FUNCTION_BLOCK MOD_StateManager (* The module's PackML state: Stopped, Resetting, Idle, Execute, Stopping, Aborted. The owner changes it with the OPC UA methods Reset, Start, Stop, Abort and Clear. It runs the Resetting and Stopping procedures and publishes the state for clients and for every block. Technical: Module state manager: OPC UA methods Reset/Start/Stop/Abort/Clear(Session) answer [Accepted, ErrorID]; publishes the PackML State over OPC UA and on the module's state channel; RUN_RESETTING and RUN_STOPPING start the procedures, which answer with *_DONE or *_FAILED *)
  (* Standard: 61499-2 *)
  (* Version 0.1, 2026-09-28, Project contributors, AAU Smart Production Lab *)
  PACKAGE modlib;
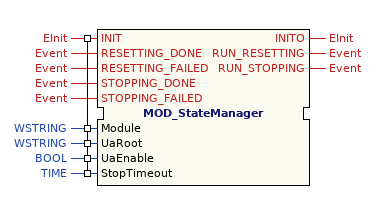
  EVENT_INPUT
    INIT : EInit WITH Module, UaRoot, UaEnable, StopTimeout; (* Initialise, once at start-up (the INIT chain); takes the values given with it *)
    RESETTING_DONE; (* The Resetting procedure ended *)
    RESETTING_FAILED; (* The Resetting procedure failed *)
    STOPPING_DONE; (* The Stopping procedure ended *)
    STOPPING_FAILED; (* The Stopping procedure failed *)
  END_EVENT
  EVENT_OUTPUT
    INITO : EInit; (* Initialised: the next block of the INIT chain goes on *)
    RUN_RESETTING; (* Run the Resetting procedure (the module was reset) *)
    RUN_STOPPING; (* Run the Stopping procedure (the module was stopped) *)
  END_EVENT
  VAR_INPUT
    Module : WSTRING; (* The module's name; its local channels are named after it (loc[<Module>/...]) *)
    UaRoot : WSTRING; (* The module's OPC UA folder, e.g. /Objects/Filling *)
    UaEnable : BOOL; (* Publish on OPC UA *)
    StopTimeout : TIME := T#10s; (* How long Stopping may take before the module aborts *)
  END_VAR
  FBS
    Ids : modlib::MOD_StateIds; (* Builds the OPC UA addresses and channel names from the module's name. *)
    Owner : modlib::MOD_OwnerView; (* Knows who occupies the module: only the owner may change the state. *)
    Reset : iec61499::net::SERVER_2_1; (* The OPC UA method Module/Reset(Session). *)
    Start : iec61499::net::SERVER_2_1; (* The OPC UA method Module/Start(Session). *)
    Stop : iec61499::net::SERVER_2_1; (* The OPC UA method Module/Stop(Session). *)
    Abort : iec61499::net::SERVER_2_1; (* The OPC UA method Module/Abort(Session). *)
    Clear : iec61499::net::SERVER_2_1; (* The OPC UA method Module/Clear(Session). *)
    Gate : modlib::MOD_StateGate; (* Decides the commands: only from the owner, only in a state PackML allows them in; answers at once. *)
    Logic : modlib::MOD_StateLogic; (* The PackML state machine. *)
    PubUa : iec61499::net::PUBLISH_1; (* Writes Module/State to OPC UA. *)
    PubState : iec61499::net::PUBLISH_1(QI := TRUE); (* Tells every block the module state, on the state channel. *)
    SubQuery : iec61499::net::SUBSCRIBE_0(QI := TRUE); (* Answers a block that asks for the state (at its start). *)
    SubAct : iec61499::net::SUBSCRIBE_1(QI := TRUE); (* Hears the skills say +1 when they start and -1 when they end. *)
    Count : modlib::MOD_ActivityCount; (* Counts the running skills: Stopping waits until none runs. *)
    Wd : iec61499::events::E_DELAY; (* Gives up waiting for the skills to stop after StopTimeout: the module then aborts. *)
  END_FBS
  EVENT_CONNECTIONS
    INIT TO Ids.INIT;
    Ids.INITO TO Owner.INIT;
    Owner.INITO TO Reset.INIT;
    Reset.INITO TO Start.INIT;
    Start.INITO TO Stop.INIT;
    Stop.INITO TO Abort.INIT;
    Abort.INITO TO Clear.INIT;
    Clear.INITO TO PubUa.INIT;
    PubUa.INITO TO PubState.INIT;
    PubState.INITO TO SubQuery.INIT;
    SubQuery.INITO TO SubAct.INIT;
    SubAct.INITO TO PubUa.REQ;
    SubAct.INITO TO PubState.REQ;
    SubAct.INITO TO INITO;
    Owner.CHG TO Gate.OWNER_CHG;
    Reset.IND TO Gate.RESET_REQ;
    Gate.RESET_RSP TO Reset.RSP;
    Gate.GO_RESET TO Logic.RESET;
    Start.IND TO Gate.START_REQ;
    Gate.START_RSP TO Start.RSP;
    Gate.GO_START TO Logic.START;
    Stop.IND TO Gate.STOP_REQ;
    Gate.STOP_RSP TO Stop.RSP;
    Gate.GO_STOP TO Logic.STOP;
    Abort.IND TO Gate.ABORT_REQ;
    Gate.ABORT_RSP TO Abort.RSP;
    Gate.GO_ABORT TO Logic.ABORT;
    Clear.IND TO Gate.CLEAR_REQ;
    Gate.CLEAR_RSP TO Clear.RSP;
    Gate.GO_CLEAR TO Logic.CLEAR;
    Logic.CNF TO PubUa.REQ;
    Logic.CNF TO PubState.REQ;
    Logic.CNF TO Gate.STATE_CHG;
    SubQuery.IND TO PubState.REQ;
    SubAct.IND TO Count.ACT;
    Count.CHG TO Logic.ACT;
    Logic.WD_START TO Wd.START;
    Logic.WD_STOP TO Wd.STOP;
    Wd.EO TO Logic.STOP_TIMEOUT;
    Logic.RUN_RESETTING TO RUN_RESETTING;
    Logic.RUN_STOPPING TO RUN_STOPPING;
    RESETTING_DONE TO Logic.RESETTING_DONE;
    RESETTING_FAILED TO Logic.RESETTING_FAILED;
    STOPPING_DONE TO Logic.STOPPING_DONE;
    STOPPING_FAILED TO Logic.STOPPING_FAILED;
  END_CONNECTIONS
  DATA_CONNECTIONS
    Module TO Ids.Module;
    Module TO Owner.Module;
    UaRoot TO Ids.UaRoot;
    UaEnable TO Reset.QI;
    UaEnable TO Start.QI;
    UaEnable TO Stop.QI;
    UaEnable TO Abort.QI;
    UaEnable TO Clear.QI;
    UaEnable TO PubUa.QI;
    StopTimeout TO Wd.DT;
    Owner.Owner TO Gate.Owner;
    Ids.IdReset TO Reset.ID;
    Reset.RD_1 TO Gate.ResetSession;
    Gate.Accepted TO Reset.SD_1;
    Gate.ErrorID TO Reset.SD_2;
    Ids.IdStart TO Start.ID;
    Start.RD_1 TO Gate.StartSession;
    Gate.Accepted TO Start.SD_1;
    Gate.ErrorID TO Start.SD_2;
    Ids.IdStop TO Stop.ID;
    Stop.RD_1 TO Gate.StopSession;
    Gate.Accepted TO Stop.SD_1;
    Gate.ErrorID TO Stop.SD_2;
    Ids.IdAbort TO Abort.ID;
    Abort.RD_1 TO Gate.AbortSession;
    Gate.Accepted TO Abort.SD_1;
    Gate.ErrorID TO Abort.SD_2;
    Ids.IdClear TO Clear.ID;
    Clear.RD_1 TO Gate.ClearSession;
    Gate.Accepted TO Clear.SD_1;
    Gate.ErrorID TO Clear.SD_2;
    Ids.IdPub TO PubUa.ID;
    Ids.IdState TO PubState.ID;
    Ids.IdQuery TO SubQuery.ID;
    Ids.IdAct TO SubAct.ID;
    Logic.State TO PubUa.SD_1;
    Logic.State TO PubState.SD_1;
    Logic.State TO Gate.State;
    SubAct.RD_1 TO Count.Delta;
    Count.AllIdle TO Logic.AllIdle;
  END_CONNECTIONS
END_FUNCTION_BLOCK
